(*
SPDX-FileCopyrightText: © 2026 Oleksandr Tiutyk <trofimich@gmail.com>
SPDX-License-Identifier: MIT
License: https://opensource.org/license/mit
*)

(*!
<summary>Checks that changing the timer preset preserves the current observation.</summary>
<description>
Starts a long interval and waits for a nonzero elapsed observation before changing the preset in RUNNING.
Also checks assignment while READY and STOPPED. One task owns the timer and AfterTest prepares it for reuse.
</description>
*)

{attribute 'no_assign'}
{attribute 'no_explicit_call' := 'do not call this function block directly'}
FUNCTION_BLOCK TimerIntervalObservationTest EXTENDS TOF_Testing.MultiCycleTest
VAR_STAT
	{attribute 'hide'}
	_ClassName : STRING := __POUNAME();
END_VAR
VAR CONSTANT
	//! <summary>Keeps the old timer active until the scenario cancels or restarts it.</summary>
	_ActiveInterval : TIME := T#1H;
END_VAR
VAR
	_Timer : TOF_Timers.Timer(name := "Configured timer");
END_VAR

(*!
<summary>Sets the initial interval while READY and starts the timer explicitly.</summary>
*)
METHOD PROTECTED BeforeTest
_Timer.Interval := _ActiveInterval;
Assert.ThatBool(
	actual := _Timer.State.Ready,
	message := "Configuring Interval must leave a READY timer idle"
).IsTrue();
Assert.ThatBool(actual := _Timer.Start(), message := "The configured timer must accept Start").IsTrue();
END_METHOD

(*!
<summary>Changes the running preset after observing positive elapsed time.</summary>
*)
METHOD PROTECTED ExecuteTest : TOF_Testing.TEST_CYCLE_RESULT
VAR
	observedTime : TIME;
END_VAR
_Timer.Execute();
observedTime := _Timer.ElapsedTime;

IF observedTime = TOF_Core.Times.MIN_VALUE THEN
	ExecuteTest := TOF_Testing.TEST_CYCLE_RESULT.BUSY;
	RETURN;
END_IF

ExecuteTest := TOF_Testing.TEST_CYCLE_RESULT.DONE;
Assert.ThatBool(
	actual := _Timer.State.Running,
	message := "A nonzero elapsed observation must belong to a running timer"
).IsTrue();
_Timer.Interval := TOF_Core.Times.MIN_VALUE;
Assert.ThatBool(
	actual := _Timer.State.Running,
	message := "Assignment of the zero preset must preserve RUNNING"
).IsTrue();
Assert.ThatBool(
	actual := _Timer.ElapsedTime = observedTime,
	message := "Assignment must preserve the nonzero elapsed observation"
).IsTrue();
Assert.ThatBool(
	actual := _Timer.Elapsed,
	message := "Assignment must leave TON.Q at its previous value"
).IsFalse();
Assert.ThatBool(
	actual := _Timer.Triggered,
	message := "Assignment must leave the completion pulse clear"
).IsFalse();

_Timer.Execute();
Assert.ThatBool(
	actual := _Timer.Triggered,
	message := "The next Execute must evaluate the changed zero preset"
).IsTrue();
observedTime := _Timer.ElapsedTime;

_Timer.Interval := _ActiveInterval;
Assert.ThatBool(
	actual := _Timer.State.Stopped,
	message := "Assigning a preset while STOPPED must keep the timer stopped"
).IsTrue();
Assert.ThatBool(
	actual := _Timer.Elapsed,
	message := "Assignment in STOPPED must preserve retained TON.Q"
).IsTrue();
Assert.ThatBool(
	actual := _Timer.ElapsedTime = observedTime,
	message := "Assignment in STOPPED must preserve elapsed time"
).IsTrue();

_Timer.Execute();
Assert.ThatBool(
	actual := _Timer.Elapsed,
	message := "Stopped Execute must preserve the retained TON observation"
).IsTrue();

IF NOT _Timer.Reset() THEN
	RecordFailure(message := "Explicit Reset must remain available after assigning the preset");
	RETURN;
END_IF

Assert.ThatBool(actual := _Timer.Elapsed, message := "Explicit Reset must clear TON.Q").IsFalse();
END_METHOD

(*!
<summary>Returns the owned timer to READY before reporting the result.</summary>
<description>
Cooperatively cancels active work and clears any retained TON observations through Reset.
</description>
*)
METHOD PROTECTED AfterTest
Assert.ThatBool(
	actual := PrepareTimerTestForReuse(timer := _Timer),
	message := "The timer must return to READY after cleanup"
).IsTrue();
END_METHOD

//! <summary>Borrows the concrete class name. Callers must not modify it.</summary>
{attribute 'monitoring' := 'call'}
PROPERTY ClassName : REFERENCE TO STRING
GET
ClassName REF= _ClassName;
END_GET
END_PROPERTY

//! <summary>Borrows the compiler-initialized namespace. Callers must not modify it.</summary>
{attribute 'monitoring' := 'call'}
PROPERTY NamespaceName : REFERENCE TO STRING
GET
NamespaceName REF= CurrentNamespace.Name;
END_GET
END_PROPERTY

//! <summary>Reports the concrete instance size in bytes.</summary>
{attribute 'monitoring' := 'call'}
PROPERTY SelfSize : ULINT
GET
SelfSize := XSIZEOF(THIS^);
END_GET
END_PROPERTY

END_FUNCTION_BLOCK

(* stored: Version 1.1.0.1
   POU TimerIntervalObservationTest: Id {89d5fbd7-c60e-4512-8015-e2b58076ca26}, SpecialFunc None
   Method BeforeTest: Id {226e26ba-e4b7-476e-9c0e-16bff1bcf052}
   Method ExecuteTest: Id {acaf479f-1e28-4ef1-ae6d-9ddc14f60cdb}
   Method AfterTest: Id {54b767a5-95a3-48f7-9f75-f28c6fd96b2f}
   Property ClassName: Id {7628572a-c3c5-401f-bc70-ae735eaf4cd5}
   Get Get: Id {c3d51b16-1795-4f42-a189-7f203d8769dd}
   Property NamespaceName: Id {61d8e1f9-83f9-4cb2-88f5-367672f00ac0}
   Get Get: Id {f942137a-f38a-487a-aa9f-69e22b50b253}
   Property SelfSize: Id {7da82b75-5b56-4490-a6f7-ce0d1e2b4e65}
   Get Get: Id {71de7b15-968d-4d80-828c-924ab4911df0} *)
